(*
SPDX-FileCopyrightText: © 2026 Oleksandr Tiutyk <trofimich@gmail.com>
SPDX-License-Identifier: MIT
License: https://opensource.org/license/mit
*)
(*!
<summary>Identifies owned directory preparation, logging, idle observation, stopping and readback phases.</summary>
*)
{attribute 'qualified_only'}
{attribute 'strict'}
TYPE LOGGER_FILE_TEST_PHASE :
(
	PREPARE_DIRECTORY,
	SEND_MESSAGES,
	OBSERVE_IDLE,
	WAIT_FOR_STOP,
	READBACK,
	COMPLETE
);
END_TYPE

(* stored: Version 1.1.0.1
   DUT LOGGER_FILE_TEST_PHASE: Id {01fb0964-31a5-4b47-9edd-30cd356f22d3} *)
